(* IEC 61131-3 sources: llm-plc-st-eval/data/processed_definitivo/claude-sonnet-4-6/A1/zero_shot, 3 files *)

(* ---- ejec_1.st ---- *)
FUNCTION_BLOCK FB_PID
VAR_INPUT
    SP    : REAL;   (* Consigna / Set Point *)
    PV    : REAL;   (* Variable de proceso *)
    Kp    : REAL;   (* Ganancia proporcional *)
    Ti    : REAL;   (* Tiempo integral [s]; <= 0 desactiva integral *)
    Td    : REAL;   (* Tiempo derivativo [s] *)
    ciclo : TIME;   (* Período de muestreo *)
END_VAR

VAR_OUTPUT
    CV : REAL;      (* Salida de mando [0.0 .. 100.0] % *)
END_VAR

VAR
    e        : REAL;   (* Error actual: SP - PV *)
    e_prev   : REAL;   (* Error en el ciclo anterior *)
    integral : REAL;   (* Acumulador de la integral del error *)
    deriv    : REAL;   (* Término derivativo *)
    Ts       : REAL;   (* Período de muestreo en segundos *)
    CV_raw   : REAL;   (* Salida sin saturar *)
    saturado : BOOL;   (* TRUE si CV está saturada *)
END_VAR

(* ── 1. Período de muestreo ─────────────────────────────────────────── *)
(* Convierte TIME → segundos; TIME_TO_DINT devuelve milisegundos *)
Ts := DINT_TO_REAL(TIME_TO_DINT(ciclo)) / 1000.0;

(* Protección: si Ts <= 0 no se puede calcular *)
IF Ts <= 0.0 THEN
    RETURN;
END_IF;

(* ── 2. Error ────────────────────────────────────────────────────────── *)
e := SP - PV;

(* ── 3. Anti-windup por clamping ─────────────────────────────────────── *)
(* Determina si la salida anterior estaba saturada *)
saturado := (CV >= 100.0) OR (CV <= 0.0);

(* Acumula integral sólo si:
   - Ti > 0  (acción integral activa)
   - No está saturado, O el error tiende a desaturar:
       · saturado en 100 → no acumular error positivo (e > 0)
       · saturado en 0   → no acumular error negativo (e < 0)       *)
IF Ti > 0.0 THEN
    IF NOT saturado
       OR (CV >= 100.0 AND e < 0.0)
       OR (CV <= 0.0  AND e > 0.0)
    THEN
        integral := integral + e * Ts;
    END_IF;
END_IF;

(* ── 4. Término derivativo ───────────────────────────────────────────── *)
deriv := (e - e_prev) / Ts;

(* ── 5. Ley de control PID (forma estándar) ──────────────────────────── *)
(*  CV = Kp · ( e  +  (1/Ti)·∫e dt  +  Td·de/dt )                       *)
IF Ti > 0.0 THEN
    CV_raw := Kp * (e + (1.0 / Ti) * integral + Td * deriv);
ELSE
    (* Sin acción integral *)
    CV_raw := Kp * (e + Td * deriv);
END_IF;

(* ── 6. Saturación de la salida ──────────────────────────────────────── *)
IF CV_raw > 100.0 THEN
    CV := 100.0;
ELSIF CV_raw < 0.0 THEN
    CV := 0.0;
ELSE
    CV := CV_raw;
END_IF;

(* ── 7. Actualiza estado para el próximo ciclo ───────────────────────── *)
e_prev := e;

END_FUNCTION_BLOCK

(* ---- ejec_2.st ---- *)
FUNCTION_BLOCK FB_PID
VAR_INPUT
    SP    : REAL;   (* Setpoint / consigna *)
    PV    : REAL;   (* Process variable / variable de proceso *)
    Kp    : REAL;   (* Ganancia proporcional *)
    Ti    : REAL;   (* Tiempo integral [s]; <= 0 desactiva integral *)
    Td    : REAL;   (* Tiempo derivativo [s] *)
    ciclo : TIME;   (* Período de muestreo *)
END_VAR

VAR_OUTPUT
    CV : REAL;      (* Salida de control [0.0 .. 100.0] % *)
END_VAR

VAR
    e_prev    : REAL;   (* Error en la iteración anterior *)
    integral  : REAL;   (* Acumulador de la integral del error *)
    Ts        : REAL;   (* Período de muestreo en segundos *)
    e         : REAL;   (* Error actual: SP - PV *)
    P_term    : REAL;   (* Término proporcional *)
    I_term    : REAL;   (* Término integral *)
    D_term    : REAL;   (* Término derivativo *)
    CV_raw    : REAL;   (* Salida sin saturar *)
    saturated : BOOL;   (* TRUE si CV está saturada *)
    sat_high  : BOOL;   (* TRUE si saturada en límite superior *)
    sat_low   : BOOL;   (* TRUE si saturada en límite inferior *)
END_VAR

(* ── Constantes de saturación ── *)
VAR CONSTANT
    CV_MAX : REAL := 100.0;
    CV_MIN : REAL := 0.0;
END_VAR

(* ─────────────────────────────────────────────────────────────
   1. Convertir período de muestreo de TIME a segundos (REAL)
   ───────────────────────────────────────────────────────────── *)
Ts := TIME_TO_REAL(ciclo) / 1000.0;   (* TIME está en ms en IEC 61131-3 *)

(* Protección: Ts debe ser positivo *)
IF Ts <= 0.0 THEN
    Ts := 0.001;   (* 1 ms mínimo para evitar división por cero *)
END_IF;

(* ─────────────────────────────────────────────────────────────
   2. Calcular error actual
   ───────────────────────────────────────────────────────────── *)
e := SP - PV;

(* ─────────────────────────────────────────────────────────────
   3. Detectar estado de saturación del ciclo anterior
   ───────────────────────────────────────────────────────────── *)
sat_high  := (CV >= CV_MAX);
sat_low   := (CV <= CV_MIN);
saturated := sat_high OR sat_low;

(* ─────────────────────────────────────────────────────────────
   4. Acumulación integral con anti-windup por clamping
      - Si saturado en máximo: no acumular error positivo
      - Si saturado en mínimo: no acumular error negativo
   ───────────────────────────────────────────────────────────── *)
IF Ti > 0.0 THEN
    IF NOT ((sat_high AND (e > 0.0)) OR (sat_low AND (e < 0.0))) THEN
        integral := integral + e * Ts;   (* Integración rectangular hacia adelante *)
    END_IF;
END_IF;

(* ─────────────────────────────────────────────────────────────
   5. Calcular términos PID
   ───────────────────────────────────────────────────────────── *)
(* Término proporcional *)
P_term := e;

(* Término integral (desactivado si Ti <= 0) *)
IF Ti > 0.0 THEN
    I_term := (1.0 / Ti) * integral;
ELSE
    I_term := 0.0;
END_IF;

(* Término derivativo: diferencia hacia atrás del error *)
D_term := Td * (e - e_prev) / Ts;

(* ─────────────────────────────────────────────────────────────
   6. Calcular salida sin saturar
   ───────────────────────────────────────────────────────────── *)
CV_raw := Kp * (P_term + I_term + D_term);

(* ─────────────────────────────────────────────────────────────
   7. Saturar salida al rango [0.0, 100.0]
   ───────────────────────────────────────────────────────────── *)
IF CV_raw >= CV_MAX THEN
    CV := CV_MAX;
ELSIF CV_raw <= CV_MIN THEN
    CV := CV_MIN;
ELSE
    CV := CV_raw;
END_IF;

(* ─────────────────────────────────────────────────────────────
   8. Guardar error para el siguiente ciclo
   ───────────────────────────────────────────────────────────── *)
e_prev := e;

(* ---- ejec_3.st ---- *)
FUNCTION_BLOCK FB_PID
VAR_INPUT
    SP    : REAL;   (* Consigna / Set Point *)
    PV    : REAL;   (* Variable de proceso / Process Variable *)
    Kp    : REAL;   (* Ganancia proporcional *)
    Ti    : REAL;   (* Tiempo integral [s]; <= 0 desactiva integral *)
    Td    : REAL;   (* Tiempo derivativo [s] *)
    ciclo : TIME;   (* Período de muestreo *)
END_VAR

VAR_OUTPUT
    CV : REAL;      (* Salida de control [0.0 .. 100.0] % *)
END_VAR

VAR
    e_prev    : REAL;   (* Error en el ciclo anterior *)
    integral  : REAL;   (* Acumulador de la integral del error *)
    dt        : REAL;   (* Período de muestreo en segundos *)
    e         : REAL;   (* Error actual: SP - PV *)
    P_term    : REAL;   (* Término proporcional *)
    I_term    : REAL;   (* Término integral *)
    D_term    : REAL;   (* Término derivativo *)
    CV_raw    : REAL;   (* Salida sin saturar *)
    saturated : BOOL;   (* TRUE si CV está saturada *)
    clamp_ok  : BOOL;   (* TRUE si se permite acumular integral *)
END_VAR

(* ── 1. Período de muestreo en segundos ─────────────────────────────── *)
dt := TIME_TO_REAL(ciclo) / 1000.0;   (* TIME está en ms en IEC 61131-3 *)

(* ── 2. Error actual ────────────────────────────────────────────────── *)
e := SP - PV;

(* ── 3. Término proporcional ────────────────────────────────────────── *)
P_term := e;

(* ── 4. Término integral con anti-windup por clamping ───────────────── *)
IF Ti > 0.0 THEN
    (* Determinar si la integración está permitida (anti-windup) *)
    (* Bloquear acumulación si CV saturada en máx y error positivo,  *)
    (* o si CV saturada en mín y error negativo.                      *)
    saturated := (CV >= 100.0) OR (CV <= 0.0);

    clamp_ok := NOT saturated                          (* sin saturación: siempre OK *)
                OR (CV >= 100.0 AND e < 0.0)          (* saturado alto, error baja  *)
                OR (CV <= 0.0  AND e > 0.0);           (* saturado bajo, error sube  *)

    IF clamp_ok THEN
        integral := integral + e * dt;
    END_IF;

    I_term := (1.0 / Ti) * integral;
ELSE
    (* Acción integral desactivada *)
    integral := 0.0;
    I_term   := 0.0;
END_IF;

(* ── 5. Término derivativo (diferencia hacia atrás sobre el error) ──── *)
IF dt > 0.0 THEN
    D_term := Td * (e - e_prev) / dt;
ELSE
    D_term := 0.0;
END_IF;

(* ── 6. Salida PID en forma estándar: CV = Kp·(e + I_term + D_term) ── *)
CV_raw := Kp * (P_term + I_term + D_term);

(* ── 7. Saturación de la salida [0.0 .. 100.0] % ───────────────────── *)
IF CV_raw > 100.0 THEN
    CV := 100.0;
ELSIF CV_raw < 0.0 THEN
    CV := 0.0;
ELSE
    CV := CV_raw;
END_IF;

(* ── 8. Guardar error para el próximo ciclo ─────────────────────────── *)
e_prev := e;

END_FUNCTION_BLOCK
